Staubli VAL3: commentIO.pgx

public program commentIO()
  local num l_i
begin

  for l_i = 0 to size(dInItem)-1
    dInItem[l_i].sComment=sCommentDin[l_i]
  endFor

  for l_i = 0 to size(dOutItem)-1
    dOutItem[l_i].sComment=sCommentDout[l_i]
  endFor

  for l_i = 0 to size(aInItem)-1
    aInItem[l_i].sComment=sCommentAin[l_i]
  endFor

  for l_i = 0 to size(aOutItem)-1
    aOutItem[l_i].sComment=sCommentAout[l_i]
  endFor

end
